(* IEC 61131-3 sources: codesys/project-view/Device/Plc Logic/Application/000-模组/本项目/00-文件读写, 5 files *)

(* ---- strFileVar.st ---- *)
TYPE strFileVar :
STRUCT

	(*文件读写变量*)
	asPara						: ARRAY[0..GlobFile.iParaLen] OF STRING;
	arNum						: ARRAY[0..GlobFile.iParaLen] OF REAL;
	asParaNum					: ARRAY[0..GlobFile.iParaLen] OF STRING;
	iFile						: UINT;
	sFileState					: STRING;//读写状态
	sFileName					: STRING:='Para_Model.txt';

END_STRUCT
END_TYPE

(* ---- uniLogPara.st ---- *)
TYPE uniLogPara :
UNION
	sLog					: STRING(GlobFile.iStringLen);
	abyLog					: ARRAY[0..GlobFile.iStringLen-1] OF BYTE;

END_UNION
END_TYPE

(* ---- GlobFile.st ---- *)
{attribute 'qualified_only'}
VAR_GLOBAL
END_VAR

VAR_GLOBAL CONSTANT
	iParaLen						: UINT:=249;//数组长度，从0开始算到iParaLen，最大值249
	iStringLen						: UINT:=20000;//文件读写的字符串总长度
// 	sNullPara						: STRING:='/ := 0.0;';//空数据连接

	sStartCharacter					: STRING:='^$R$N';//起始符
	sTerminator						: STRING:='#';//终止符

END_VAR

(* ---- FUN_ReadFileArray.st ---- *)
//读取文件，将字符串里的数据分成数组[0..199]
//数据完整返回'OK'，否则返回'NG'
FUNCTION FUN_ReadFileArray : STRING
VAR_INPUT
	FilePath						: STRING;
END_VAR

VAR_OUTPUT
	sReceData						: STRING(GlobFile.iStringLen);				//读取的字符串(无处理)
	asParaNum						: ARRAY[0..GlobFile.iParaLen] OF STRING;	//读取分割后的数据字符串数组
	arNum							: ARRAY[0..GlobFile.iParaLen] OF REAL;		//读取的数据
END_VAR

VAR
	i								: UINT;
	uniLogPara						: uniLogPara;

	FileHandle						: RTS_IEC_HANDLE;
	ResError1						: RTS_IEC_RESULT;
	ResError2						: RTS_IEC_RESULT;
	ResError3						: RTS_IEC_RESULT;

	sIsComplete						: STRING;//字符串是否完整
	iFind							: ARRAY[0..1] OF INT;
	asTmp							: ARRAY[0..GlobFile.iParaLen] OF STRING;

END_VAR

VAR CONSTANT
	sConnect						: STRING:='$R$N';

END_VAR
// --- implementation ---
(**************************************************************
例如：
sReceData := '123$R$N456';

输出：
arNum[0] => 123;			arNum[1] => 456;

***************************************************************)

// //清除数据
// sReceData := '';
// FOR i:=0 TO GlobFile.iParaLen DO
// 	arNum[i] := 0;
// END_FOR

//打开文件
FileHandle:= SysFileOpen(szFile:= FilePath, am:= ACCESS_MODE.AM_READ_PLUS, pResult:= ADR(ResError1));

//读取数据
SysFileRead(hFile:= FileHandle, pbyBuffer:= ADR(uniLogPara.abyLog[0]), ulSize:=SIZEOF(uniLogPara.abyLog), pResult:=ADR(ResError2));

//关闭文件
SysFileClose(hFile:= FileHandle);

sReceData := uniLogPara.sLog;

(*********************************		处理字符串		*********************************)

//检查字符串是否完整
sIsComplete := FUN_CheckString(RcvStr:=uniLogPara.sLog , StartStr:=GlobFile.sStartCharacter , EndStr:=GlobFile.sTerminator , xFromStr=>uniLogPara.sLog );

IF sIsComplete = 'OK' THEN	//数据完整

	//将字符串分割成字符串数组
	FUN_CutString(sString:=uniLogPara.sLog , sStartCharacter:='/' , sTerminator:=';' , asParaNum=>asParaNum );

	//提取字符串数组' := '后面的数据
	FOR i := 0 TO GlobFile.iParaLen DO
		IF asParaNum[i] = '' THEN//空数据，跳出循环
			EXIT;
		ELSE
			arNum[i] := TO_REAL(	FUN_FindString(str:=asParaNum[i] , str1:=':= ' , str2:=';' )	);

		END_IF

	END_FOR

	FUN_ReadFileArray := 'OK';

ELSE	//数据不完整，报错

	FUN_ReadFileArray := 'NG';

END_IF

(******************************************************
//此部分是预留，如果字符串长度超过255，可以使用此部分

iFind[0] := FIND(STR1:=asParaNum[i] , STR2:=':= ' );		//查询':= '的位置
iFind[1] := FIND(STR1:=asParaNum[i] , STR2:=';' );			//查询';'的位置
StrMidA(
	pst := ADR(asParaNum[i]),
	uiInputBufferSize := SIZEOF(ADR(asParaNum[i])),
	iLength := iFind[1] - iFind[0] - len(':= '), 		//计算提取数据的长度。从':= '开始数，到';'结束，其中还要减去':= '自身长度
	iPosition := iFind[0] + len(':= '), 				//从':= '最右边开始提取，所以加上':= '自身长度
	pstResult := ADR(asTmp[i]),
	uiResultBufferSize := 0);
arNum[i] := TO_REAL(asTmp[i]);

**********************************************************)
END_FUNCTION

(* ---- FUN_WriteFileArray.st ---- *)
//将字符串数组[0..199]中每个元素合并，以'$R$N'连接，并写入文件
FUNCTION FUN_WriteFileArray : STRING
VAR_INPUT
	FilePath						: STRING;
	asParaNum						: ARRAY[0..GlobFile.iParaLen] OF STRING;
END_VAR

VAR
	uniLogPara						: uniLogPara;//写入文件的字符串
	i								: UINT;
	sTmp							: STRING(GlobFile.iStringLen);

	FileHandle						: RTS_IEC_HANDLE;
	ResError1						: RTS_IEC_RESULT;
	ResError2						: RTS_IEC_RESULT;
	ResError3						: RTS_IEC_RESULT;

END_VAR

VAR CONSTANT
	sConnect						: STRING:='$R$N';
// 	sStart							: STRING(GlobFile.iStringLen):='^$R$N';
// 	sFinal							: STRING:='#';
END_VAR
// --- implementation ---
(**************************************************************
数组元素合并
例如：
asParaNum[0] := '123';			asParaNum[1] := '456';

输出：
sParaWtrie => '123$R$N456';

***************************************************************)

(*****************	处理字符串，使之与上面注释描述连接	**********************)

FOR i := 0 TO TO_UINT(GlobFile.iParaLen) DO

	//如果这个数据是空数据，就跳出循环，不连接空数据
	IF asParaNum[i] = '' THEN//GlobFile.sNullPara THEN
		EXIT;
	END_IF

	//连接字符串
	IF i = 0 THEN
		uniLogPara.sLog := CONCAT(STR1:=GlobFile.sStartCharacter , STR2:=asParaNum[i] );//最前面加个'^$R$N'作起始符号
		StrConcatA(pstFrom:=ADR(sConnect) , pstTo:=ADR(uniLogPara.sLog) , iBufferSize:=TO_INT(SIZEOF(uniLogPara.sLog)) );
	ELSE
		StrConcatA(pstFrom:=ADR(asParaNum[i]) , pstTo:=ADR(uniLogPara.sLog) , iBufferSize:=TO_INT(SIZEOF(uniLogPara.sLog)) );
		StrConcatA(pstFrom:=ADR(sConnect) , pstTo:=ADR(uniLogPara.sLog) , iBufferSize:=TO_INT(SIZEOF(uniLogPara.sLog)) );

	END_IF

END_FOR

//最后加个'#'作结束符号
StrConcatA(pstFrom:=ADR(GlobFile.sTerminator) , pstTo:=ADR(uniLogPara.sLog) , iBufferSize:=TO_INT(SIZEOF(uniLogPara.sLog)) );

(***********************************************************************************************)

//为了避免写入数据长度出错的问题，先删除文件，再写入
// SysFileDeleteByHandle(hFile:=FileHandle );
SM3_Basic.SysFileDelete(szFileName:=FilePath );

//打开文件
FileHandle:= SysFileOpen(szFile:= FilePath, am:= ACCESS_MODE.AM_WRITE_PLUS, pResult:= ADR(ResError1));

//设置写入的偏移位置，每次都从第一个位置开始复写
// SysFileSetPos(hFile:= FileHandle, ulOffset:=SysFileGetSize(szFileName:= FilePath, pResult:= ADR(ResError2)) );

//写入数据
SM3_Basic.SysFileWrite(hFile:= FileHandle, pbyBuffer:= ADR(uniLogPara.abyLog), ulSize:= TO_LWORD(StrLenA(pstData:=ADR(uniLogPara.sLog)) ), pResult:= ADR(ResError3));

//关闭文件
SysFileClose(hFile:= FileHandle);
END_FUNCTION
